       REGION 正常状态判断
           IF NOT "v_bianliang".dianti[#i].cuowu.REP_deal AND NOT "v_bianliang".dianti[#i].Weight_handle.jiangyao_chaozhong AND NOT "v_bianliang".dianti[#i].Weight_handle.chaozhongxinhao THEN
               "v_bianliang".dianti[#i].报警指示灯 := 1;
           END_IF;

       END_REGION

       IF "IO".elev[#i].jinggao.REP OR "v_bianliang".dianti[#i].cuowu.qi_ting THEN
           "v_bianliang".dianti[#i].cuowu.REP_deal := 1;
       ELSE                                                   
           "v_bianliang".dianti[#i].cuowu.REP_deal := 0;
       END_IF;
       //检修处理
       IF "v_bianliang".dianti[#i].cuowu.REP_deal THEN
           "报警".维修报警[#i] := 1;
           "v_bianliang".dianti[#i].状态指示灯 := 2;
           "v_bianliang".dianti[#i].报警指示灯 := 3;
           "IO".elev[#i].display.error := 1; //亮起故障指示灯
           // IF "v_bianliang".dianti[#i].interrupt.f_100ms = 1 THEN
           //     "v_bianliang".dianti[#i].interrupt.f_100ms := 0;
           //     CASE "v_bianliang".dianti[#i].interrupt.state OF
           //         0:

           //             "v_bianliang".dianti[#i].interrupt.state := 1;
           //         1:
           //             "IO".elev[#i].display.error := 0;
           //             "v_bianliang".dianti[#i].interrupt.state := 0;
           //     END_CASE;
           // END_IF;
               "v_bianliang".dianti[#i].yunxing_chuli.yunxu_run := 0; //该电梯停止运行
               "v_bianliang".dianti[#i].init.kaishi := 0;//不进行初始化

               "v_bianliang".dianti[#i].yunxing_chuli.run_state := 0; //运行状态机为静止态
               "v_bianliang".dianti[#i].yunxing_chuli.uopdown_state := 0; //上下行状态为静止
               //电梯控制状态为静止:关闭电机、接触器
               "run_state"(eet_num := #i,
                           state :="STATIC");
       END_IF;
       //检测检修信号下降沿:检测到下降沿，电梯进行初始化后投入使用
       IF NOT "v_bianliang".dianti[#i].cuowu.REP_deal AND "v_bianliang".dianti[#i].cuowu.tag_REPL THEN //若检测到下降沿
           "v_bianliang".dianti[#i].init.kaishi := 1;//让该部电梯开始初始化
           "IO".elev[#i].display.error := 0; //关闭故障指示灯
           "报警".维修报警[#i] := 0;

           IF "v_bianliang".dianti[#i].init.re_mode =1 THEN //手动设置检修后初始化方向
               "v_bianliang".dianti[#i].init.init_fangxiang := "v_bianliang".dianti[#i].init.re_fangxiang;
               IF "v_bianliang".dianti[#i].init.re_fangxiang THEN //向上初始化停在10层
                   "v_bianliang".dianti[#i].init.mubiao_floor := "FlOOR_TOP";
               ELSE
                   "v_bianliang".dianti[#i].init.mubiao_floor := 1;
               END_IF;
           ELSIF "v_bianliang".dianti[#i].Floor_handle.dangqian_floor = 0 THEN //若该电梯当前楼层为0，则说明在初始化前该电梯就开始检修
               "v_bianliang".dianti[#i].init.init_fangxiang := "v_bianliang".dianti[#i].gaibian.init_dir; //初始化方向就为预设方向
               IF NOT "v_bianliang".dianti[#i].gaibian.init_dir THEN //下行撞限位就停到1层
                   "v_bianliang".dianti[#i].init.mubiao_floor := 1;
               ELSE
                   "v_bianliang".dianti[#i].init.mubiao_floor := "FlOOR_TOP";//否则停到十层
               END_IF;
           ELSE //若该电梯有楼层，则说明是在运行时检修的，那么则就近初始化
               IF "v_bianliang".dianti[#i].Floor_handle.dangqian_floor <= 5 THEN //楼层在5层即以下，向下初始化停在一层
                   "v_bianliang".dianti[#i].init.init_fangxiang := 0;
                   "v_bianliang".dianti[#i].init.mubiao_floor := 1;
               ELSE //否则向上初始化停到10层
                   "v_bianliang".dianti[#i].init.init_fangxiang := 1;
                   "v_bianliang".dianti[#i].init.mubiao_floor := "FlOOR_TOP";
               END_IF;
           END_IF;
       END_IF;
       "v_bianliang".dianti[#i].cuowu.tag_REPL := "v_bianliang".dianti[#i].cuowu.REP_deal; //将检修信号存入tag中 
   END_FOR;
END_FUNCTION

FUNCTION "Weight_judgement" : Void   // FC12, SCL
{ S7_Optimized_Access := 'TRUE' }
VERSION : 0.1
   VAR_TEMP
      i : Int;
   END_VAR
BEGIN

   FOR #i := 1 TO "ELE_SUM" DO
       "v_bianliang".dianti[#i].Weight_handle.m_load := NORM_X(MIN := 0, VALUE := "IO".elev[#i].zhongliang, MAX := 27648);
       "v_bianliang".dianti[#i].Weight_handle.shiji_load := SCALE_X(MIN := 0, VALUE := "v_bianliang".dianti[#i].Weight_handle.m_load, MAX := 2000);
   END_FOR;


   FOR #i := 1 TO "ELE_SUM" DO
       "v_bianliang".dianti[#i].Weight_handle.max_load := "v_bianliang".dianti[#i].gaibian.max_load;
   END_FOR;


   FOR #i := 1 TO "ELE_SUM" DO 
       IF ("v_bianliang".dianti[#i].Weight_handle.shiji_load  > "v_bianliang".dianti[#i].Weight_handle.max_load) OR "v_bianliang".dianti[#i].gaibian.now_load> "v_bianliang".dianti[#i].Weight_handle.max_load THEN
           "v_bianliang".dianti[#i].Weight_handle.chaozhongxinhao := 1;

           IF "v_bianliang".dianti[#i].yunxing_chuli.uopdown_state = 1 THEN//该电梯在该楼层超载，该楼层的外呼信号直接分配给群控，不要等外呼按钮
               "v_bianliang".anniu_waibu[1, "v_bianliang".dianti[#i].Floor_handle.dangqian_floor] := 1;
           ELSIF "v_bianliang".dianti[#i].yunxing_chuli.uopdown_state = 2 THEN
               "v_bianliang".anniu_waibu[2, "v_bianliang".dianti[#i].Floor_handle.dangqian_floor] := 1;
           END_IF;

           "报警".超重报警[#i] := 1;
           "v_bianliang".dianti[#i].报警指示灯 := 4;
       ELSE
           "v_bianliang".dianti[#i].Weight_handle.chaozhongxinhao := 0;
           "报警".超重报警[#i] := 0;
       END_IF;


       IF ("v_bianliang".dianti[#i].Weight_handle.shiji_load > "v_bianliang".dianti[#i].Weight_handle.max_load - 75) OR "v_bianliang".dianti[#i].gaibian.now_load > "v_bianliang".dianti[#i].Weight_handle.max_load - 75 THEN
           "v_bianliang".dianti[#i].Weight_handle.jiangyao_chaozhong := 1;
       ELSE
           "v_bianliang".dianti[#i].Weight_handle.jiangyao_chaozhong := 0;
       END_IF;

       IF "v_bianliang".dianti[#i].Weight_handle.jiangyao_chaozhong = 1 AND NOT "v_bianliang".dianti[#i].Weight_handle.chaozhongxinhao THEN
           "v_bianliang".dianti[#i].状态指示灯 := 2;
           "v_bianliang".dianti[#i].报警指示灯 := 2;
       END_IF;

   END_FOR;
END_FUNCTION

FUNCTION "RUN_CTL_ALL" : Void   // FC13, SCL
{ S7_Optimized_Access := 'TRUE' }
VERSION : 0.1
   VAR_TEMP
      i : Int;
      j : Int;
      start : Bool;
   END_VAR
BEGIN
   FOR #i := 1 TO "ELE_SUM" DO
       IF "v_bianliang".dianti[#i].yunxing_chuli.yunxu_run THEN

           "select_updown"(i := #i);

           CASE "v_bianliang".dianti[#i].yunxing_chuli.run_state OF
               0:
                   REGION 初始态，电梯由静止转向运动
                       "run_state"(eet_num := #i,
                                        state := "STATIC");//静止

                       IF "v_bianliang".dianti[#i].yunxing_chuli.uopdown_state = 1 AND NOT "IO".elev[#i].direction.up AND "IO".elev[#i].direction.down THEN
                           "v_bianliang".dianti[#i].Count[3].CV := "v_bianliang".dianti[#i].Count[3].CV + 1;
                       ELSIF "v_bianliang".dianti[#i].yunxing_chuli.uopdown_state = 2 AND "IO".elev[#i].direction.up AND NOT "IO".elev[#i].direction.down THEN
                           "v_bianliang".dianti[#i].Count[3].CV := "v_bianliang".dianti[#i].Count[3].CV - 1;
                       END_IF;

                       IF "v_bianliang".dianti[#i].yunxing_chuli.uopdown_state = 1 THEN
                           "v_bianliang".dianti[#i].yunxing_chuli.run_state := 1;
                       ELSIF "v_bianliang".dianti[#i].yunxing_chuli.uopdown_state = 2 THEN 
                           "v_bianliang".dianti[#i].yunxing_chuli.run_state := 2;
                       ELSIF "v_bianliang".dianti[#i].yunxing_chuli.uopdown_state = 0 THEN 
                           "v_bianliang".dianti[#i].yunxing_chuli.run_state := 0;
                       END_IF;

                       IF ("v_bianliang".dianti[#i].yunxing_chuli.uopdown_state = 1 AND "v_bianliang".dianti[#i].anniu_luru.waibu_anniu[1, "v_bianliang".dianti[#i].Floor_handle.dangqian_floor]) OR
                           ("v_bianliang".dianti[#i].yunxing_chuli.uopdown_state = 2 AND "v_bianliang".dianti[#i].anniu_luru.waibu_anniu[2, "v_bianliang".dianti[#i].Floor_handle.dangqian_floor]) AND
                           "IO".elev[#i].direction.up AND "IO".elev[#i].direction.down THEN 
                           "v_bianliang".dianti[#i].yunxing_chuli.run_state := 6;
                       END_IF;
                   END_REGION
               1:
                   REGION 上行启动态，低速启动
                       "run_state"(eet_num := #i,
                                        state := "UP_L"); 

                       "v_bianliang".dianti[#i].shijian[1].TON(IN := "IO".elev[#i].ele_speed.L,
                                                 PT := T#0.1S);
                       IF "v_bianliang".dianti[#i].shijian[1].Q THEN 
                           "v_bianliang".dianti[#i].yunxing_chuli.run_state := 3;
                       END_IF;
                   END_REGION
               2:
                   REGION 下行启动态，低速启动
                       "run_state"(eet_num := #i,
                                       state := "DOWN_L"); 

                       "v_bianliang".dianti[#i].shijian[1].TON(IN := "IO".elev[#i].ele_speed.L,
                                                 PT := T#0.1S);
                       IF "v_bianliang".dianti[#i].shijian[1].Q THEN 
                           "v_bianliang".dianti[#i].yunxing_chuli.run_state := 4;
                       END_IF;
                   END_REGION
               3:
                   REGION 上行态
                       "run_state"(eet_num := #i,
                                       state := "UP_H");//上行高速

                       IF ("v_bianliang".dianti[#i].yunxing_chuli.uopdown_state = 0 OR "v_bianliang".dianti[#i].yunxing_chuli.uopdown_state = 2)
                           AND "IO".elev[#i].direction.up THEN 
                           "v_bianliang".dianti[#i].yunxing_chuli.run_state := 5;
                       END_IF;

                       IF "v_bianliang".dianti[#i].Weight_handle.jiangyao_chaozhong THEN //将超载时只响应内呼
                           IF "v_bianliang".dianti[#i].anniu_luru.neibu_anniu["v_bianliang".dianti[#i].Floor_handle.dangqian_floor] AND "IO".elev[#i].direction.up THEN
                               "v_bianliang".dianti[#i].yunxing_chuli.run_state := 5;
                           END_IF;
                       ELSE //正常响应
                           IF (("v_bianliang".dianti[#i].anniu_luru.waibu_anniu[1, "v_bianliang".dianti[#i].Floor_handle.dangqian_floor] OR "v_bianliang".dianti[#i].anniu_luru.neibu_anniu["v_bianliang".dianti[#i].Floor_handle.dangqian_floor])
                               OR ("v_bianliang".dianti[#i].Floor_handle.dangqian_floor = "v_bianliang".dianti[#i].yunxing_chuli.zuida_floor AND "v_bianliang".dianti[#i].anniu_luru.waibu_anniu[2, "v_bianliang".dianti[#i].yunxing_chuli.zuida_floor]))
                               AND "IO".elev[#i].direction.up AND NOT "IO".elev[#i].direction.down THEN
                               "v_bianliang".dianti[#i].yunxing_chuli.run_state := 5;
                           ELSIF "v_bianliang".dianti[#i].Floor_handle.dangqian_floor=10 AND "IO".elev[#i].direction.up AND NOT "IO".elev[#i].direction.down THEN//若到十层，强制制动
                               "v_bianliang".dianti[#i].yunxing_chuli.run_state := 5;
                           END_IF;
                       END_IF;
                   END_REGION
               4:
                   REGION 下行态
                       "run_state"(eet_num := #i,
                                       state := "DOWN_H"); 

                       IF ("v_bianliang".dianti[#i].yunxing_chuli.uopdown_state = 0 OR "v_bianliang".dianti[#i].yunxing_chuli.uopdown_state = 1)
                           AND "IO".elev[#i].direction.down THEN 
                           "v_bianliang".dianti[#i].yunxing_chuli.run_state := 5;
                       END_IF;

                       IF "v_bianliang".dianti[#i].Weight_handle.jiangyao_chaozhong THEN 
                           IF "v_bianliang".dianti[#i].anniu_luru.neibu_anniu["v_bianliang".dianti[#i].Floor_handle.dangqian_floor] AND "IO".elev[#i].direction.down THEN
                               "v_bianliang".dianti[#i].yunxing_chuli.run_state := 5;
                           END_IF;
                       ELSE //正常响应
                           IF (("v_bianliang".dianti[#i].anniu_luru.waibu_anniu[2, "v_bianliang".dianti[#i].Floor_handle.dangqian_floor] OR "v_bianliang".dianti[#i].anniu_luru.neibu_anniu["v_bianliang".dianti[#i].Floor_handle.dangqian_floor])
                               OR ("v_bianliang".dianti[#i].Floor_handle.dangqian_floor = "v_bianliang".dianti[#i].yunxing_chuli.zuixiao_floor AND "v_bianliang".dianti[#i].anniu_luru.waibu_anniu[1, "v_bianliang".dianti[#i].yunxing_chuli.zuixiao_floor]))
                               AND "IO".elev[#i].direction.down AND NOT "IO".elev[#i].direction.up THEN
                               "v_bianliang".dianti[#i].yunxing_chuli.run_state := 5;
                           ELSIF "v_bianliang".dianti[#i].Floor_handle.dangqian_floor=1 AND NOT "IO".elev[#i].direction.up AND "IO".elev[#i].direction.down THEN//若到一层，强制制动
                               "v_bianliang".dianti[#i].yunxing_chuli.run_state := 5;
                           END_IF;
                       END_IF;
                   END_REGION
               5:
                   REGION 减速制动态 ，电梯到达指定楼层减速制动     
                       IF "v_bianliang".dianti[#i].gaibian.speed = 1 THEN 
                           IF "IO".elev[#i].direction.down AND "IO".elev[#i].direction.up THEN 
                               "run_state"(eet_num := #i,
                                               state := "H_L"); 
                           END_IF;
                           "v_bianliang".dianti[#i].shijian[3].TON(IN := "IO".elev[#i].ele_speed.L,
                                                     PT := T#1MS,
                                                     Q => "IO".elev[#i].Brake.B1);
                           "v_bianliang".dianti[#i].shijian[4].TON(IN := "IO".elev[#i].Brake.B1,
                                                     PT := T#1MS,
                                                     Q => "IO".elev[#i].Brake.B2);
                           "v_bianliang".dianti[#i].shijian[5].TON(IN := "IO".elev[#i].Brake.B2,
                                                     PT := T#1MS,
                                                     Q => "IO".elev[#i].Brake.B3);
                       ELSIF "v_bianliang".dianti[#i].gaibian.speed = 2 THEN //中速电梯制动
                           #start := 1; //启动定时器的标志变量
                           "v_bianliang".dianti[#i].shijian[2].TON(IN := #start, //延迟一段时间转低速制动
                                                     PT := T#0.4S);
                           IF "v_bianliang".dianti[#i].shijian[2].Q THEN
                               "run_state"(eet_num := #i,
                                               state := "H_L");//高速转低速
                           END_IF;
                           "v_bianliang".dianti[#i].shijian[3].TON(IN := "IO".elev[#i].ele_speed.L,
                                                     PT := T#0.7S,
                                                     Q => "IO".elev[#i].Brake.B1);
                           "v_bianliang".dianti[#i].shijian[4].TON(IN := "IO".elev[#i].Brake.B1,
                                                     PT := T#1MS,
                                                     Q => "IO".elev[#i].Brake.B2);
                           "v_bianliang".dianti[#i].shijian[5].TON(IN := "IO".elev[#i].Brake.B2,
                                                     PT := T#1MS,
                                                     Q => "IO".elev[#i].Brake.B3);
                       ELSIF "v_bianliang".dianti[#i].gaibian.speed = 3 THEN //高速电梯制动
                           #start := 1; //启动定时器的标志变量
                           "v_bianliang".dianti[#i].shijian[2].TON(IN := #start, //延迟一段时间转低速制动
                                                     PT := T#0.25S);
                           IF "v_bianliang".dianti[#i].shijian[2].Q THEN
                               "run_state"(eet_num := #i,
                                               state := "H_L");
                           END_IF;
                           "v_bianliang".dianti[#i].shijian[3].TON(IN := "IO".elev[#i].ele_speed.L,
                                                     PT := T#1MS,
                                                     Q => "IO".elev[#i].Brake.B1);
                           "v_bianliang".dianti[#i].shijian[4].TON(IN := "IO".elev[#i].Brake.B1,
                                                     PT := T#1MS,
                                                     Q => "IO".elev[#i].Brake.B2);
                           "v_bianliang".dianti[#i].shijian[5].TON(IN := "IO".elev[#i].Brake.B2,
                                                     PT := T#1MS,
                                                     Q => "IO".elev[#i].Brake.B3);
                       END_IF;
                       IF "IO".elev[#i].Brake.B3 THEN
                           //正常转消层态
                           "v_bianliang".dianti[#i].yunxing_chuli.run_state := 6;

                       END_IF;
                   END_REGION
               6:
                   REGION 消层态，当电梯到达目标楼层后，消除内外呼信号
                       "run_state"(eet_num := #i,
                                       state := "STATIC"); //静止

                       RESET_TIMER("v_bianliang".dianti[#i].shijian[1]);
                       RESET_TIMER("v_bianliang".dianti[#i].shijian[2]);
                       RESET_TIMER("v_bianliang".dianti[#i].shijian[3]);
                       RESET_TIMER("v_bianliang".dianti[#i].shijian[4]);
                       RESET_TIMER("v_bianliang".dianti[#i].shijian[5]);

                       "IO".elev[#i].Brake.B1 := 0;
                       "IO".elev[#i].Brake.B2 := 0;
                       "IO".elev[#i].Brake.B3 := 0;

                       "v_bianliang".dianti[#i].anniu_luru.neibu_anniu["v_bianliang".dianti[#i].Floor_handle.dangqian_floor] := 0;

                       IF "v_bianliang".dianti[#i].yunxing_chuli.uopdown_state = 1 THEN //若是上行 则消除上呼
                           "v_bianliang".anniu_waibu[1, "v_bianliang".dianti[#i].Floor_handle.dangqian_floor] := 0;
                           "v_bianliang".dianti[#i].anniu_luru.waibu_anniu[1, "v_bianliang".dianti[#i].Floor_handle.dangqian_floor] := 0;
                           "v_bianliang".flag[1] := 1;

                       ELSIF "v_bianliang".dianti[#i].yunxing_chuli.uopdown_state = 2 THEN//若是下行 则消除下呼
                           "v_bianliang".dianti[#i].anniu_luru.waibu_anniu[2, "v_bianliang".dianti[#i].Floor_handle.dangqian_floor] := 0;
                           "v_bianliang".anniu_waibu[2, "v_bianliang".dianti[#i].Floor_handle.dangqian_floor] := 0;
                           "v_bianliang".flag[2] := 1;

                       END_IF;

                       "v_bianliang".dianti[#i].yunxing_chuli.run_state := 7;
                   END_REGION
               7:
                   REGION 消层后，电梯开门
                       "run_state"(eet_num := #i,
                                       state := "OPEN");
                           "v_bianliang".dianti[#i].shijian[6].TON(IN := "IO".elev[#i].door_jdq.open,
                                                                   PT := T#4.4S);

                         IF "v_bianliang".dianti[#i].shijian[6].Q THEN
                             "v_bianliang".dianti[#i].yunxing_chuli.run_state := 8;
                         END_IF;
                   END_REGION
               8:
                   REGION 开门后，电梯关门
                       RESET_TIMER("v_bianliang".dianti[#i].shijian[6]);
                       IF "IO".elev[#i].door_inplace.close = 0 AND "IO".elev[#i].jinggao.LC = 0 AND "v_bianliang".dianti[#i].Weight_handle.chaozhongxinhao = 0 THEN
                           "run_state"(eet_num := #i,
                                           state := "CLOSE");
                       END_IF;
                       IF "IO".elev[#i].door_inplace.close = 0 AND ("IO".elev[#i].jinggao.LC = 1 OR "v_bianliang".dianti[#i].Weight_handle.chaozhongxinhao = 1) THEN
                           "run_state"(eet_num := #i,
                                       state := "OPEN");
                           "v_bianliang".dianti[#i].shijian[12].TON(IN := "IO".elev[#i].door_inplace.close = 0,
                                                      PT := T#120MS);
                           IF "v_bianliang".dianti[#i].shijian[12].Q THEN
                               "v_bianliang".dianti[#i].yunxing_chuli.run_state := 8;
                               RESET_TIMER("v_bianliang".dianti[#i].shijian[12]);
                           END_IF;
                       END_IF;

                       IF "IO".elev[#i].door_inplace.close THEN
                           "v_bianliang".dianti[#i].yunxing_chuli.run_state := 0;

                           IF "v_bianliang".flag[1] = 1 THEN
                               "v_bianliang".flag[1] := 0;
                               "v_bianliang".start_tim[1, "v_bianliang".dianti[#i].Floor_handle.dangqian_floor] := "v_bianliang".all_time.min * 60 + "v_bianliang".all_time.sec;//开始的时间
                           ELSIF "v_bianliang".flag[2] = 1 THEN
                               "v_bianliang".flag[2] := 0;
                               "v_bianliang".start_tim[2, "v_bianliang".dianti[#i].Floor_handle.dangqian_floor] := "v_bianliang".all_time.min * 60 + "v_bianliang".all_time.sec;//开始的时间
                           END_IF;

                       END_IF;

                       //若不在将超载时，有人按下本层外呼，
                       IF NOT "v_bianliang".dianti[#i].Weight_handle.jiangyao_chaozhong THEN
                           IF "v_bianliang".dianti[#i].yunxing_chuli.uopdown_state = 1 THEN //若是上行 则消除上呼
                               "v_bianliang".anniu_waibu[1, "v_bianliang".dianti[#i].Floor_handle.dangqian_floor] := 0;
                               "v_bianliang".dianti[#i].anniu_luru.waibu_anniu[1, "v_bianliang".dianti[#i].Floor_handle.dangqian_floor] := 0;
                           ELSIF "v_bianliang".dianti[#i].yunxing_chuli.uopdown_state = 2 THEN//若是下行 则消除下呼
                               "v_bianliang".dianti[#i].anniu_luru.waibu_anniu[2, "v_bianliang".dianti[#i].Floor_handle.dangqian_floor] := 0;
                               "v_bianliang".anniu_waibu[2, "v_bianliang".dianti[#i].Floor_handle.dangqian_floor] := 0;
                           END_IF;
                       END_IF;
                   END_REGION
               9:
                   REGION 超重处理态
                       "run_state"(eet_num := #i,
                                       state := "OPEN");

                       IF NOT "v_bianliang".dianti[#i].Weight_handle.chaozhongxinhao THEN
                           "v_bianliang".dianti[#i].yunxing_chuli.run_state := 8;
                       END_IF;
                   END_REGION ;       
           END_CASE;
       END_IF;

       IF "v_bianliang".dianti[#i].yunxing_chuli.yunxu_run THEN
           "v_bianliang".dianti[#i].状态指示灯 := 1;
       END_IF;
   END_FOR;
END_FUNCTION

FUNCTION "select_updown" : Void   // FC14, SCL
{ S7_Optimized_Access := 'TRUE' }
VERSION : 0.1
   VAR_INPUT
      i : Int;
   END_VAR
   VAR_TEMP
      j : Int;
      p : Bool;
      q : Bool;
   END_VAR
BEGIN
   "v_bianliang".dianti[#i].yunxing_chuli.zuida_floor := 0; //判断最高层
   IF "v_bianliang".dianti[#i].yunxing_chuli.uopdown_state <> 2 AND "v_bianliang".dianti[#i].Floor_handle.dangqian_floor <> 0 THEN //电梯不下行时，判断最高层
       FOR #j := "v_bianliang".dianti[#i].Floor_handle.dangqian_floor TO "FlOOR_TOP"  DO //判断当前层到最高层
           IF "v_bianliang".dianti[#i].anniu_luru.waibu_anniu[1, #j] OR "v_bianliang".dianti[#i].anniu_luru.neibu_anniu[#j] OR "v_bianliang".dianti[#i].anniu_luru.waibu_anniu[2, #j] THEN
               "v_bianliang".dianti[#i].yunxing_chuli.zuida_floor := #j;
           END_IF;
       END_FOR;
   END_IF;

   "v_bianliang".dianti[#i].yunxing_chuli.zuixiao_floor  := 0;//判断最底层
   IF "v_bianliang".dianti[#i].yunxing_chuli.uopdown_state <> 1 AND "v_bianliang".dianti[#i].Floor_handle.dangqian_floor<>0 THEN//电梯不上行，判断最底层
       FOR #j := "v_bianliang".dianti[#i].Floor_handle.dangqian_floor TO 1 BY -1 DO //判断当前楼层到最底层
           IF "v_bianliang".dianti[#i].anniu_luru.waibu_anniu[2, #j] OR "v_bianliang".dianti[#i].anniu_luru.neibu_anniu[#j] OR "v_bianliang".dianti[#i].anniu_luru.waibu_anniu[1, #j] THEN
               "v_bianliang".dianti[#i].yunxing_chuli.zuixiao_floor := #j;
           END_IF;
       END_FOR;
   END_IF;
   //判断运行方向
   IF "v_bianliang".dianti[#i].yunxing_chuli.zuida_floor  > "v_bianliang".dianti[#i].Floor_handle.dangqian_floor THEN //先判断上方，若存在最高层，先向上运行
       "v_bianliang".dianti[#i].yunxing_chuli.uopdown_state := 1;
   ELSIF "v_bianliang".dianti[#i].yunxing_chuli.zuida_floor  = "v_bianliang".dianti[#i].Floor_handle.dangqian_floor THEN //到达最高层后,判断继续向上还是转向
       IF "v_bianliang".dianti[#i].anniu_luru.waibu_anniu[1, "v_bianliang".dianti[#i].Floor_handle.dangqian_floor ] THEN //若最远层是上呼，那么则继续上行
           "v_bianliang".dianti[#i].yunxing_chuli.uopdown_state := 1;
       ELSIF "v_bianliang".dianti[#i].anniu_luru.waibu_anniu[2, "v_bianliang".dianti[#i].Floor_handle.dangqian_floor ] THEN //若最远层是下呼，那么则转向
           "v_bianliang".dianti[#i].yunxing_chuli.uopdown_state := 2;
       ELSE
           "v_bianliang".dianti[#i].yunxing_chuli.uopdown_state := 0;//最远层是内呼则静止
       END_IF;
   END_IF;

   IF "v_bianliang".dianti[#i].yunxing_chuli.zuixiao_floor < "v_bianliang".dianti[#i].Floor_handle.dangqian_floor AND "v_bianliang".dianti[#i].yunxing_chuli.zuixiao_floor <> 0 THEN //先判断下方，若存在最低层，先向下运行
       "v_bianliang".dianti[#i].yunxing_chuli.uopdown_state := 2;
   ELSIF "v_bianliang".dianti[#i].yunxing_chuli.zuixiao_floor = "v_bianliang".dianti[#i].Floor_handle.dangqian_floor THEN //到达最低层后，判断继续向下还是转向
       IF "v_bianliang".dianti[#i].anniu_luru.waibu_anniu[2, "v_bianliang".dianti[#i].Floor_handle.dangqian_floor] THEN //若最远层是下呼，那么则继续下行
           "v_bianliang".dianti[#i].yunxing_chuli.uopdown_state := 2;
       ELSIF "v_bianliang".dianti[#i].anniu_luru.waibu_anniu[1, "v_bianliang".dianti[#i].Floor_handle.dangqian_floor] THEN //若最远层是上呼，那么则转向
           "v_bianliang".dianti[#i].yunxing_chuli.uopdown_state := 1;
       ELSE
           "v_bianliang".dianti[#i].yunxing_chuli.uopdown_state := 0;//最远层是内呼则静止
       END_IF;
   END_IF;

   //最底层和最高层间强制转向
   IF "v_bianliang".dianti[#i].yunxing_chuli.run_state <> 0 THEN
       IF "v_bianliang".dianti[#i].Floor_handle.dangqian_floor = 1 THEN //在一层强制上行
           "v_bianliang".dianti[#i].yunxing_chuli.uopdown_state := 1;
       ELSIF "v_bianliang".dianti[#i].Floor_handle.dangqian_floor = 10 THEN //在十层强制下行
           "v_bianliang".dianti[#i].yunxing_chuli.uopdown_state := 2;
       END_IF;
   END_IF;
   //判断静止状态
   IF "v_bianliang".dianti[#i].yunxing_chuli.run_state = 8 AND "IO".elev[#i].door_inplace.close THEN //若电梯开门后又关门且关门完毕
       IF ("v_bianliang".dianti[#i].yunxing_chuli.zuida_floor = 0 AND "v_bianliang".dianti[#i].yunxing_chuli.uopdown_state = 1) OR//若上行但无最高层
           ("v_bianliang".dianti[#i].yunxing_chuli.zuixiao_floor = 0 AND "v_bianliang".dianti[#i].yunxing_chuli.uopdown_state = 2) THEN //或下行但无最低层
           "v_bianliang".dianti[#i].yunxing_chuli.uopdown_state := 0; //则电梯静止
       END_IF;
   END_IF;
END_FUNCTION

FUNCTION "nei_hu" : Void   // FC15, SCL
{ S7_Optimized_Access := 'TRUE' }
VERSION : 0.1
   VAR_INPUT
      i : Int;
      j : Int;
   END_VAR
BEGIN
   IF "IO".elev[#i].ele_in_button[#j].state AND NOT "IO".elev[#i].ele_in_button[#j].p THEN
       //正向登陆
       IF "v_bianliang".dianti[#i].yunxing_chuli.uopdown_state = 0 OR
           ("v_bianliang".dianti[#i].yunxing_chuli.uopdown_state = 1 AND #j > "v_bianliang".dianti[#i].Floor_handle.dangqian_floor) OR
           ("v_bianliang".dianti[#i].yunxing_chuli.uopdown_state = 2 AND #j < "v_bianliang".dianti[#i].Floor_handle.dangqian_floor) THEN
           "v_bianliang".dianti[#i].anniu_luru.neibu_anniu[#j] := 1;
           "IO".elev[#i].ele_in_button[#j].light := 1;
           //反向登陆    
       ELSIF ("v_bianliang".dianti[#i].yunxing_chuli.uopdown_state = 1 AND #j < "v_bianliang".dianti[#i].Floor_handle.dangqian_floor) OR
           ("v_bianliang".dianti[#i].yunxing_chuli.uopdown_state = 2 AND #j > "v_bianliang".dianti[#i].Floor_handle.dangqian_floor) THEN
           "v_bianliang".dianti[#i].anniu_luru.neibu_anniu[#j] := 1;
       END_IF;
   END_IF;

   "IO".elev[#i].ele_in_button[#j].p := "IO".elev[#i].ele_in_button[#j].state;

   IF "v_bianliang".dianti[#i].anniu_luru.neibu_anniu[#j] = 0 THEN
       "IO".elev[#i].ele_in_button[#j].light := 0;
   END_IF;
END_FUNCTION

FUNCTION "GP_CTL" : Void   // FC16, SCL
{ S7_Optimized_Access := 'TRUE' }
VERSION : 0.1
   VAR_TEMP
      i : Int;
      j : Int;
      p : Bool;
      q : Bool;
   END_VAR
BEGIN
   FOR #j := 1 TO "FlOOR_TOP" DO 
       REGION 当前楼层外呼分配
           FOR #i := 1 TO "ELE_SUM" DO
               IF "v_bianliang".dianti[#i].yunxing_chuli.uopdown_state = 0 AND "v_bianliang".dianti[#i].cuowu.REP_deal = 0 THEN
                   IF "v_bianliang".anniu_waibu[1, "v_bianliang".dianti[#i].Floor_handle.dangqian_floor] AND "v_bianliang".dianti[#i].Floor_handle.dangqian_floor = #j THEN
                       "v_bianliang"."dianti"[#i].anniu_luru.waibu_anniu[1, #j] := 1;
                   ELSIF "v_bianliang".anniu_waibu[2, "v_bianliang".dianti[#i].Floor_handle.dangqian_floor] AND "v_bianliang".dianti[#i].Floor_handle.dangqian_floor = #j THEN
                       "v_bianliang"."dianti"[#i].anniu_luru.waibu_anniu[2, #j] := 1;
                   END_IF;
                   EXIT;
               END_IF;
           END_FOR;
       END_REGION

       REGION 该层有无分配信号判断
           #p := 0;//该层上呼判断
           #q := 0;//该层下呼判断
           FOR #i := 1 TO "ELE_SUM" DO
               IF "v_bianliang".dianti[#i].anniu_luru.waibu_anniu[1, #j] THEN 
                   #p := 1;
               END_IF;
               IF "v_bianliang".dianti[#i].anniu_luru.waibu_anniu[2, #j] THEN 
                   #q := 1;
               END_IF;
           END_FOR;
           IF (NOT "v_bianliang".anniu_waibu[1, #j] AND NOT "v_bianliang".anniu_waibu[2, #j]) OR (#p AND #q) THEN
               CONTINUE;
           END_IF;
       END_REGION

       REGION 清空时间计算
           FOR #i := 1 TO "ELE_SUM" DO
               "v_bianliang".dianti[#i].qunkong.TH := 0;
           END_FOR;
       END_REGION

       REGION 上呼梯信号时间计算
           FOR #i := 1 TO "ELE_SUM" DO
               IF "v_bianliang".anniu_waibu[1, #j] AND NOT #p AND "v_bianliang".dianti[#i].Floor_handle.dangqian_floor <> #j THEN //判断是否有上呼且该层上呼没有被分配
                   "count_staytime"(VC := "v_bianliang".dianti[#i].yunxing_chuli.uopdown_state, //传入电梯当前运行方向
                                  F0 := "v_bianliang".dianti[#i].Floor_handle.dangqian_floor,       //传入电梯当前楼层
                                  V := "v_bianliang".dianti[#i].gaibian.speed,            //传入电梯当前速度
                                  X := #i,                                     //传入当前电梯序列
                                  FS := #j,                                    //传入当前处理的楼层
                                  VA := 1);                                    //传入外呼方向：1上
               END_IF;
           END_FOR;
       END_REGION

       REGION 上呼梯信号分配
           IF "v_bianliang".anniu_waibu[1, #j] AND NOT #p THEN
               "compare_tim"();
               "desperate_task"(aim_f := #j);
               IF "v_bianliang".zuiyou_dianti <> 0 THEN
                   "v_bianliang"."dianti"["v_bianliang".zuiyou_dianti].anniu_luru.waibu_anniu[1, #j] := 1;//分配给上呼内信号

               END_IF;
           END_IF;
       END_REGION

       REGION 清空时间计算
           FOR #i := 1 TO "ELE_SUM" DO
               "v_bianliang".dianti[#i].qunkong.TH := 0;
           END_FOR;
       END_REGION

       REGION 下呼梯信号时间计算
           FOR #i := 1 TO "ELE_SUM" DO
               IF "v_bianliang".anniu_waibu[2, #j] AND NOT #q AND "v_bianliang".dianti[#i].Floor_handle.dangqian_floor <> #j THEN //判断是否有下呼且该层下呼没有被分配
                   "count_staytime"(VC := "v_bianliang".dianti[#i].yunxing_chuli.uopdown_state, //传入电梯当前运行方向
                                  F0 := "v_bianliang".dianti[#i].Floor_handle.dangqian_floor,       //传入电梯当前楼层
                                  V := "v_bianliang".dianti[#i].gaibian.speed,            //传入电梯当前速度
                                  X := #i,                                     //传入当前电梯序列
                                  FS := #j,                                    //传入当前处理的楼层
                                  VA := 2);                                    //传入外呼方向：2下
                END_IF;
           END_FOR;
       END_REGION

       REGION 下呼梯信号分配
           IF "v_bianliang".anniu_waibu[2, #j] AND NOT #p THEN
               "compare_tim"();
               "desperate_task"(aim_f := #j);
               IF "v_bianliang".zuiyou_dianti <> 0 THEN 
                   "v_bianliang".dianti["v_bianliang".zuiyou_dianti].anniu_luru.waibu_anniu[2, #j] := 1; //分配给下呼内信号
               END_IF;

           END_IF; 
       END_REGION
   END_FOR;
   "clear_mission"();
END_FUNCTION

FUNCTION "count_staytime" : Void   // FC17, SCL
{ S7_Optimized_Access := 'TRUE' }
VERSION : 0.1
   VAR_INPUT
      VC : Int;   // 电梯运行方向
      F0 : Int;   // 当前楼层
      V : Int;   // 电梯速度
      X : Int;   // 当前处理电梯
      FS : Int;   // 处理楼层
      VA : Int;   // 外呼呼叫方向
   END_VAR
   VAR_TEMP
      i : Int;
      Fmax : Int;   // 同向运行最远楼层
      Fmin : Int;   // 反向运行最远楼层
      TD : Int;   // 经过一个楼层时间
      TK : Int;   // 停层时间
      N : Int;   // 任务数
   END_VAR
BEGIN
   REGION 参数设定     
       CASE #V OF
           1://低速
               #TD := 67; 
               #TK := 130;   
           2: //中速
               #TD := 40;
               #TK := 130; 
           3://高速
               #TD := 27; 
               #TK := 130; 
       END_CASE;
   END_REGION


   CASE #VC OF
       0:
           REGION 电梯静止时
               "v_bianliang".dianti[#X].qunkong.TH := ABS(#FS - #F0) * #TD; //候梯时间即为层差
           END_REGION
       1:
           REGION 电梯上行时
               IF #VA = 1 THEN 
                   IF #FS >= #F0 THEN 
                       #N := 0;
                       FOR #i := #F0 TO #FS DO 
                           IF "v_bianliang".dianti[#X].anniu_luru.neibu_anniu[#i] OR "v_bianliang".dianti[#X].anniu_luru.waibu_anniu[1, #i] THEN
                               #N += 1;
                           END_IF;
                       END_FOR;
                       "v_bianliang".dianti[#X].qunkong.TH := ABS(#FS - #F0) * #TD + #N * #TK; 
                   ELSE
                       "v_bianliang".dianti[#X].qunkong.TH := 10000;
                   END_IF;
               ELSIF #VA = 2 THEN 
                   FOR #i := #F0 TO 1 BY -1 DO 
                       IF "v_bianliang".dianti[#X].anniu_luru.neibu_anniu[#i] OR "v_bianliang".dianti[#X].anniu_luru.waibu_anniu[2, #i] THEN
                           #Fmin := #i;
                       END_IF;
                   END_FOR;
                   #N := 0;
                   FOR #i := #F0 TO #Fmin DO 
                       IF "v_bianliang".dianti[#X].anniu_luru.neibu_anniu[#i] OR "v_bianliang".dianti[#X].anniu_luru.waibu_anniu[1, #i] OR "v_bianliang".dianti[#X].anniu_luru.waibu_anniu[2, #i] THEN
                           #N += 1;
                       END_IF;
                   END_FOR;
                   "v_bianliang".dianti[#X].qunkong.TH := ABS(#Fmin - #F0) * #TD + ABS(#FS - #Fmin) * #TD + #N * #TK + #TD;
               END_IF;
           END_REGION
       2:
           REGION 电梯下行时
               IF #VA = 2 THEN //信号为下呼，只考虑下呼在下方，在后方的下呼默认时间最久
                   IF #FS <= #F0 THEN //当呼梯信号在本层或下方
                       #N := 0;//任务数清0
                       FOR #i := #FS TO #F0 DO //计算任务数
                           IF "v_bianliang".dianti[#X].anniu_luru.neibu_anniu[#i] OR "v_bianliang".dianti[#X].anniu_luru.waibu_anniu[2, #i] THEN
                               #N += 1;
                           END_IF;
                       END_FOR;
                       "v_bianliang".dianti[#X].qunkong.TH := ABS(#FS - #F0) * #TD + #N * #TK; //侯梯时间等于电梯经过楼层时间+停层时间
                   ELSE
                       "v_bianliang".dianti[#X].qunkong.TH := 10000;
                   END_IF;
               ELSIF #VA = 1 THEN //信号为上呼
                   FOR #i := #F0 TO "FlOOR_TOP" DO //计算上行最远层
                       IF "v_bianliang".dianti[#X].anniu_luru.neibu_anniu[#i] OR "v_bianliang".dianti[#X].anniu_luru.waibu_anniu[1, #i] THEN
                           #Fmax := #i;
                       END_IF;
                   END_FOR;
                   #N := 0;//任务数清0
                   FOR #i := #F0 TO #Fmax DO //计算任务数
                       IF "v_bianliang".dianti[#X].anniu_luru.neibu_anniu[#i] OR "v_bianliang".dianti[#X].anniu_luru.waibu_anniu[1, #i] OR "v_bianliang".dianti[#X].anniu_luru.waibu_anniu[2, #i] THEN
                           #N += 1;
                       END_IF;
                   END_FOR;
                   "v_bianliang".dianti[#X].qunkong.TH := ABS(#Fmin - #F0) * #TD + ABS(#FS - #Fmin) * #TD + #N * #TK +#TD;//候梯时间为电梯到最小层再折回到呼梯楼层+停层时间
               END_IF;
           END_REGION
   END_CASE;
   IF NOT "v_bianliang".dianti[#X].yunxing_chuli.yunxu_run THEN 
       "v_bianliang".dianti[#X].qunkong.TH := 10000;
   END_IF;

   IF "v_bianliang".dianti[#X].Weight_handle.jiangyao_chaozhong AND NOT "v_bianliang".dianti[#X].anniu_luru.neibu_anniu[#FS] THEN 
       "v_bianliang".dianti[#X].qunkong.TH := 10000;
   END_IF;

   // REGION 分区的补丁
   //     IF #FS = 2 AND #X <> 5 THEN//除了5号梯，其他的电梯都不去2楼
   //         "v_bianliang".dianti[#X].qunkong.TH := 10000;
   //     END_IF;

   //     IF (#FS = 3 OR #FS = 4) AND #X = 6 THEN
   //         "v_bianliang".dianti[#X].qunkong.TH := 10000;
   //     END_IF;
   // END_REGION


   // IF "variable".elevator[#X].Weight_handle.to_overload THEN//将要超载不响应外呼
   //     "variable".elevator[#X].group_control.TH := 10000;
   // END_IF;

   // "variable".elevator[#i].Weight_handle.now_load > "variable".elevator[#i].Weight_handle.max_load - 75 #FS = 1 OR #FS = 3 OR #FS = 5 OR #FS = 7 OR #FS = 9 THEN
   //     "variable".elevator[1].group_control.TH := 10000;
   //     "variable".elevator[3].group_control.TH := 10000;
   // END_IF;

   // IF #FS = 2 OR #FS = 3 OR #FS = 4 OR #FS = 5 OR #FS = 6 AND NOT "variable".elevator[1].Btn_Input.inside[#FS] THEN
   //     "variable".elevator[1].group_control.TH := 10000;
   // END_IF;

   // IF #FS = 2  OR #FS = 6 AND NOT "variable".elevator[2].Btn_Input.inside[#FS] THEN
   //     "variable".elevator[2].group_control.TH := 10000;
   // END_IF;


   // 
   // IF "variable".elevator[1].Weight_handle.now_load > "variable".elevator[1].Weight_handle.max_load - 75 * 2 THEN
   //     "variable".elevator[1].group_control.TH := 10000;
   // END_IF;
   //
END_FUNCTION

FUNCTION "compare_tim" : Void   // FC18, SCL
{ S7_Optimized_Access := 'TRUE' }
VERSION : 0.1
   VAR_TEMP
      i : Int;
      j : Int;
      temp : Int;
      temp_num : Int;
   END_VAR
BEGIN

   FOR #i := 1 TO "ELE_SUM" DO 
       "v_bianliang".time_min[#i] := #i;
   END_FOR;

   FOR #i := 1 TO "ELE_SUM" DO
       IF "v_bianliang".dianti[#i].qunkong.TH = 0 THEN
           "v_bianliang".dianti[#i].qunkong.TH := 10000;
       END_IF;
   END_FOR;

   FOR #i := 1 TO "ELE_SUM" DO
           FOR #j := 1 TO "ELE_SUM" - #i DO
               IF "v_bianliang".dianti[#j].qunkong.TH > "v_bianliang".dianti[#j + 1].qunkong.TH THEN 
                   #temp := "v_bianliang".dianti[#j].qunkong.TH;
                   "v_bianliang".dianti[#j].qunkong.TH := "v_bianliang".dianti[#j + 1].qunkong.TH;
                   "v_bianliang".dianti[#j + 1].qunkong.TH := #temp;

                   #temp_num := "v_bianliang".time_min[#j];        
                   "v_bianliang".time_min[#j] := "v_bianliang".time_min[#j + 1];
                   "v_bianliang".time_min[#j + 1] := #temp_num;
               END_IF;
           END_FOR;
   END_FOR;
END_FUNCTION

FUNCTION "desperate_task" : Void   // FC19, SCL
{ S7_Optimized_Access := 'TRUE' }
VERSION : 0.1
   VAR_INPUT
      aim_f : Int;
   END_VAR
   VAR_TEMP
      i : Int;
      j : Int;
      temp : Int;
      flag : Bool;
   END_VAR
BEGIN
   FOR #i := 1 TO "ELE_SUM" DO
       IF "v_bianliang".dianti[#i].qunkong.TH < 500 THEN 
           EXIT;
       ELSE 
           "v_bianliang".zuiyou_dianti := 0;
           RETURN;
       END_IF;
   END_FOR;

   FOR #i := 1 TO "ELE_SUM" DO
       IF "v_bianliang".dianti[#i].Weight_handle.chaozhongxinhao THEN
           IF "v_bianliang".dianti[#i].yunxing_chuli.uopdown_state = 1 THEN
               "v_bianliang".anniu_waibu[1, "v_bianliang".dianti[#i].Floor_handle.dangqian_floor] := 1;
           ELSIF "v_bianliang".dianti[#i].yunxing_chuli.uopdown_state = 2 THEN 
               "v_bianliang".anniu_waibu[2, "v_bianliang".dianti[#i].Floor_handle.dangqian_floor] := 1;
           END_IF;
       END_IF;
   END_FOR;


   "v_bianliang".zuiyou_dianti := "v_bianliang".time_min[1];
END_FUNCTION

FUNCTION "clear_mission" : Void   // FC20, SCL
{ S7_Optimized_Access := 'TRUE' }
VERSION : 0.1
   VAR_TEMP
      i : Int;
      j : Int;
      k : Int;
      cnt_tag : Int;
      tag : Bool;
      flag_up : Bool;
      flag_down : Bool;
   END_VAR
BEGIN
   //若外呼消除，
   FOR #j := 2 TO "FlOOR_TOP" -1 DO
       FOR #i := 1 TO "ELE_SUM" DO
           IF NOT "v_bianliang".anniu_waibu[1, #j] THEN
               "v_bianliang".dianti[#i].anniu_luru.waibu_anniu[1, #j] := 0;
           END_IF;
           IF NOT "v_bianliang".anniu_waibu[2, #j] THEN
               "v_bianliang".dianti[#i].anniu_luru.waibu_anniu[2, #j] := 0;
           END_IF;
       END_FOR;
   END_FOR;
   //当一部电梯将要超载时，
   FOR #i := 1 TO "ELE_SUM" DO
       IF "v_bianliang".dianti[#i].Weight_handle.jiangyao_chaozhong THEN
           FOR #j := 1 TO "FlOOR_TOP" DO
               IF ("v_bianliang".dianti[#i].anniu_luru.waibu_anniu[1, #j] OR "v_bianliang".dianti[#i].anniu_luru.waibu_anniu[2, #j]) AND NOT "v_bianliang".dianti[#i].anniu_luru.neibu_anniu[#j] THEN
                   "v_bianliang".dianti[#i].anniu_luru.waibu_anniu[1, #j] := 0;
                   "v_bianliang".dianti[#i].anniu_luru.waibu_anniu[2, #j] := 0;
               END_IF;
           END_FOR;
       END_IF;
   END_FOR;
   //当电梯检修时
   FOR #i := 1 TO "ELE_SUM" DO
       IF NOT "v_bianliang".dianti[#i].yunxing_chuli.yunxu_run THEN
           FOR #j := 1 TO "FlOOR_TOP" DO
               "v_bianliang".dianti[#i].anniu_luru.waibu_anniu[1, #j] := 0;
               "v_bianliang".dianti[#i].anniu_luru.waibu_anniu[2, #j] := 0;
           END_FOR;
       END_IF;
   END_FOR;
   //清除电梯的后方外呼
   FOR #i := 1 TO "ELE_SUM" DO
       IF "v_bianliang".dianti[#i].yunxing_chuli.uopdown_state = 1 AND "v_bianliang".dianti[#i].Floor_handle.dangqian_floor>1 THEN
           FOR #j := 1 TO "v_bianliang".dianti[#i].Floor_handle.dangqian_floor - 1 DO
               "v_bianliang".dianti[#i].anniu_luru.waibu_anniu[1, #j] := 0;
               "v_bianliang".dianti[#i].anniu_luru.waibu_anniu[2, #j] := 0;
           END_FOR;
       ELSIF "v_bianliang".dianti[#i].yunxing_chuli.uopdown_state = 2 AND "v_bianliang".dianti[#i].Floor_handle.dangqian_floor<"FlOOR_TOP" THEN
           FOR #j := "FlOOR_TOP" TO "v_bianliang".dianti[#i].Floor_handle.dangqian_floor + 1 BY -1 DO
               "v_bianliang".dianti[#i].anniu_luru.waibu_anniu[1, #j] := 0;
               "v_bianliang".dianti[#i].anniu_luru.waibu_anniu[2, #j] := 0;
           END_FOR;
       END_IF;
   END_FOR;
   //若一部电梯没有任务
   FOR #i := 1 TO "ELE_SUM" DO
       IF "v_bianliang".dianti[#i].yunxing_chuli.uopdown_state = 0 AND "v_bianliang".dianti[#i].yunxing_chuli.yunxu_run THEN
           #tag := 1;
           EXIT;
       END_IF;
       IF "v_bianliang".dianti[#i].yunxing_chuli.uopdown_state <> 0 OR NOT "v_bianliang".dianti[#i].yunxing_chuli.yunxu_run THEN
           #cnt_tag += 1;
       END_IF;
   END_FOR;
   IF #cnt_tag = "ELE_SUM" THEN
       #tag := 0;
   END_IF;
   "R_TRIG_DB"(CLK:=#tag);
   IF "R_TRIG_DB".Q THEN
       FOR #i := 1 TO "ELE_SUM" DO
           FOR #j := 1 TO "FlOOR_TOP" DO
               IF #j <> "v_bianliang".dianti[#i].Floor_handle.dangqian_floor THEN
                   "v_bianliang".dianti[#i].anniu_luru.waibu_anniu[1, #j] := 0;
                   "v_bianliang".dianti[#i].anniu_luru.waibu_anniu[2, #j] := 0;
               END_IF;
           END_FOR;
       END_FOR;
   END_IF;


   //优先响应最优上呼
   FOR #i := 1 TO "ELE_SUM" DO
       IF "v_bianliang"."dianti"[#i].anniu_luru.waibu_anniu[1, "v_bianliang".zuiyou_louceng[1]] AND "v_bianliang".slope[1, "v_bianliang".zuiyou_louceng[1]] > 70 THEN
           FOR #j := 1 TO "FlOOR_TOP" - 1 DO
               IF "v_bianliang".zuiyou_louceng[1] <> #j THEN//除了最优呼梯，其他呼梯都不响应
                   "v_bianliang".dianti[#i].anniu_luru.waibu_anniu[1, #j] := 0;
               END_IF;
           END_FOR;
           EXIT;
       END_IF;
   END_FOR;

   //优先响应最优下呼
   FOR #i := 1 TO "ELE_SUM" DO
       IF "v_bianliang"."dianti"[#i].anniu_luru.waibu_anniu[2, "v_bianliang".zuiyou_louceng[2]] AND "v_bianliang".slope[2, "v_bianliang".zuiyou_louceng[2]] > 70 THEN
           FOR #j := 2 TO "FlOOR_TOP" DO
               IF "v_bianliang".zuiyou_louceng[2] <> #j THEN//除了最优呼梯，其他呼梯都不响应
                   "v_bianliang".dianti[#i].anniu_luru.waibu_anniu[2, #j] := 0;
               END_IF;
           END_FOR;
           EXIT;
       END_IF;
   END_FOR;


   // FOR #i := 2 TO "ELE_SUM" DO //早高峰的补丁，当3号到6号梯没有任务且是允许运行的时候，该电梯停在一楼
   //     IF "v_bianliang".dianti[#i].yunxing_chuli.uopdown_state = 0 AND "v_bianliang".dianti[#i].yunxing_chuli.yunxu_run THEN
   //         "v_bianliang".dianti[#i].anniu_luru.neibu_anniu[7] := 1;
   //         IF "v_bianliang".dianti[#i].Floor_handle.dangqian_floor = 7 THEN
   //             "v_bianliang".dianti[#i].anniu_luru.neibu_anniu[7] := 0;
   //         END_IF;
   //     END_IF;
   // END_FOR;

   // //若执行同向任务时又接收反向任务，则将距离>1的反向任务清除
   // FOR #i := 1 TO "ELE_SUM" DO
   //     #flag_up := 0;
   //     FOR #j := 1 TO "FlOOR_TOP" DO
   //         IF "Var".elev[#i].Run_Deal.uopdown_state = 1 AND "Var".elev[#i].Btn_Input.outside[1, #j] THEN
   //             #flag_up := 1;
   //             GOTO LABEL1;
   //         ELSE
   //             EXIT;
   //         END_IF;
   //     END_FOR;
   //     LABEL1:
   //     IF #flag_up THEN
   //         FOR #j := 1 TO "FlOOR_TOP" DO
   //             IF #j <> "Var".elev[#i].Floor_Deal.Now_f THEN
   //                 "Var".elev[#i].Btn_Input.outside[2, #j] := 0;
   //             END_IF;
   //         END_FOR;
   //     END_IF;

   //     #flag_down := 0;
   //     FOR #j := 1 TO "FlOOR_TOP" DO
   //         IF "Var".elev[#i].Run_Deal.uopdown_state = 2 AND "Var".elev[#i].Btn_Input.outside[2, #j] THEN
   //             #flag_down := 1;
   //             GOTO LABEL2;
   //         ELSE
   //             EXIT;
   //         END_IF;
   //     END_FOR;
   //     LABEL2:
   //     IF #flag_down THEN
   //         FOR #j := 1 TO "FlOOR_TOP" DO
   //             IF #j <> "Var".elev[#i].Floor_Deal.Now_f THEN
   //                 "Var".elev[#i].Btn_Input.outside[1, #j] := 0;
   //             END_IF;
   //         END_FOR;
   //     END_IF;
   // END_FOR;
END_FUNCTION

FUNCTION "Guard" : Void   // FC21, SCL
{ S7_Optimized_Access := 'TRUE' }
VERSION : 0.1
   VAR_TEMP
      i : Int;
   END_VAR
BEGIN
   FOR #i := 1 TO "ELE_SUM" DO
       IF "v_bianliang".dianti[#i].yunxing_chuli.yunxu_run THEN
           IF "IO".elev[#i].bt_limit.bottom1 AND "v_bianliang".dianti[#i].yunxing_chuli.run_state = 4 THEN
               "v_bianliang".dianti[#i].yunxing_chuli.run_state := 3;
               "v_bianliang".dianti[#i].yunxing_chuli.uopdown_state := 1;
               "v_bianliang".dianti[#i].Count[3].CV := 1;
           ELSIF "IO".elev[#i].bt_limit.top1 AND "v_bianliang".dianti[#i].yunxing_chuli.run_state = 3 THEN
               "v_bianliang".dianti[#i].yunxing_chuli.run_state := 4;
               "v_bianliang".dianti[#i].yunxing_chuli.uopdown_state := 2;
               "v_bianliang".dianti[#i].Count[3].CV := 10;
           END_IF;
       END_IF;
   END_FOR;
END_FUNCTION

FUNCTION "forecast" : Void   // FC22, SCL
{ S7_Optimized_Access := 'TRUE' }
VERSION : 0.1
   VAR_TEMP
      i : Int;
      j : Int;
      temp : Real;
      flour_temp : Int;
      max : Real;
   END_VAR
BEGIN
   FOR #i := 1 TO "ELE_SUM" DO
       FOR #j := 1 TO "FlOOR_TOP" DO
           IF "v_bianliang".over_tim[1, #j] > "v_bianliang".start_tim[1, #j] AND "v_bianliang".dianti[#i].Floor_handle.dangqian_floor = #j THEN//结束时间<开始时间且有电梯再此楼层，标志位加一
               "v_bianliang".dianti[#i].flag[1, #j] := 1;
           END_IF;

           IF ("v_bianliang".start_tim[1, #j] < ("v_bianliang".all_time.min * 60 + "v_bianliang".all_time.sec)) AND "v_bianliang".dianti[#i].flag[1, #j] = 1 THEN
               "v_bianliang".dianti[#i].flag[1, #j] := 0;
               #temp:=("v_bianliang".over_tim[1, #j] - "v_bianliang".start_tim[1, #j]);//转化浮点数类型
               "v_bianliang".slope[1, #j] :=  "v_bianliang".dianti[#i].Weight_handle.shiji_load*1.0/#temp ;
           END_IF;

           IF "v_bianliang".over_tim[2, #j] > "v_bianliang".start_tim[2, #j] AND "v_bianliang".dianti[#i].Floor_handle.dangqian_floor = #j THEN//结束时间<开始时间且有电梯再此楼层，标志位加一
               "v_bianliang".dianti[#i].flag[2, #j] := 1;
           END_IF;

           IF ("v_bianliang".start_tim[2, #j] < ("v_bianliang".all_time.min * 60 + "v_bianliang".all_time.sec)) AND "v_bianliang".dianti[#i].flag[2, #j] = 1 THEN
               "v_bianliang".dianti[#i].flag[2, #j] := 0;
               #temp:=("v_bianliang".over_tim[2, #j] - "v_bianliang".start_tim[2, #j]);//转化浮点数类型
               "v_bianliang".slope[2, #j] :=  "v_bianliang".dianti[#i].Weight_handle.shiji_load*1.0/#temp ;
           END_IF;
       END_FOR;
   END_FOR;

   #max := "v_bianliang".slope[1, 1];//判断最优上呼楼层

   FOR #j := 1 TO "FlOOR_TOP"-1 DO
       IF "v_bianliang".slope[1, #j] >= #max THEN
           #max := "v_bianliang".slope[1, #j];
           "v_bianliang".zuiyou_louceng[1] := #j;
       END_IF;
   END_FOR;

   #max := "v_bianliang".slope[2, 2];//判断最优下呼楼层

   FOR #j := 2 TO "FlOOR_TOP"DO
       IF "v_bianliang".slope[2, #j] >= #max THEN
           #max := "v_bianliang".slope[2, #j];
           "v_bianliang".zuiyou_louceng[2] := #j;
       END_IF;
   END_FOR;
END_FUNCTION

ORGANIZATION_BLOCK "Main"   // OB1, LAD, ProgramCycle
TITLE = "Main Program Sweep (Cycle)"
{ S7_Optimized_Access := 'TRUE' }
VERSION : 0.1
   VAR_INPUT
      Initial_Call : Bool;   // Initial call of this OB
      Remanence : Bool;   // =True, if remanent data are available
   END_VAR
BEGIN

REGION Network 1 (SCL)
   "addr management"();                   

   "init_signal"();                        
   "signal_check"();                        
   "init_up"();                           
   // "timer"();                      //定时器

   IF "IO".plc_ready THEN

   "show_F"();                         
   "CALL_ELE"();                           
   "Weight_judgement"();
   "forecast"();//预测
   "GP_CTL"();                      
   "RUN_CTL_ALL"();                      
   "Indicate"();                         
   "Guard"();

   END_IF;
END_REGION
END_ORGANIZATION_BLOCK

ORGANIZATION_BLOCK "Cyclic interrupt"   // OB30, LAD, CyclicInterrupt
{ S7_Optimized_Access := 'TRUE' }
VERSION : 0.1
   VAR_INPUT
      Initial_Call : Bool;   // Initial call of this OB
      Event_Count : Int;   // Events discarded
   END_VAR
   VAR_TEMP
      i : Int;
      cnt_1s : Int;
   END_VAR
BEGIN

REGION Network 1 (SCL)

   // FOR #i :=1 TO "ELE_SUM" DO
   //     "v_bianliang".dianti[#i].interrupt.f_1ms:= 1;
   // END_FOR;

   IF "IO".plc_ready THEN
       "v_bianliang".all_time.cnt_1s += 1;
       IF "v_bianliang".all_time.cnt_1s > 999 THEN
           "v_bianliang".all_time.cnt_1s := 0;
           "v_bianliang".all_time.sec += 1;
       END_IF;
       IF "v_bianliang".all_time.sec > 59 THEN
           "v_bianliang".all_time.sec := 0;
           "v_bianliang".all_time.min += 1;
       END_IF;
       IF "v_bianliang".all_time.min > 59 THEN
           "v_bianliang".all_time.min := 0;
           "v_bianliang".all_time.hour += 1;
       END_IF;
       IF "v_bianliang".all_time.hour > 23 THEN
           "v_bianliang".all_time.hour := 0;
       END_IF;
   END_IF;
END_REGION
END_ORGANIZATION_BLOCK